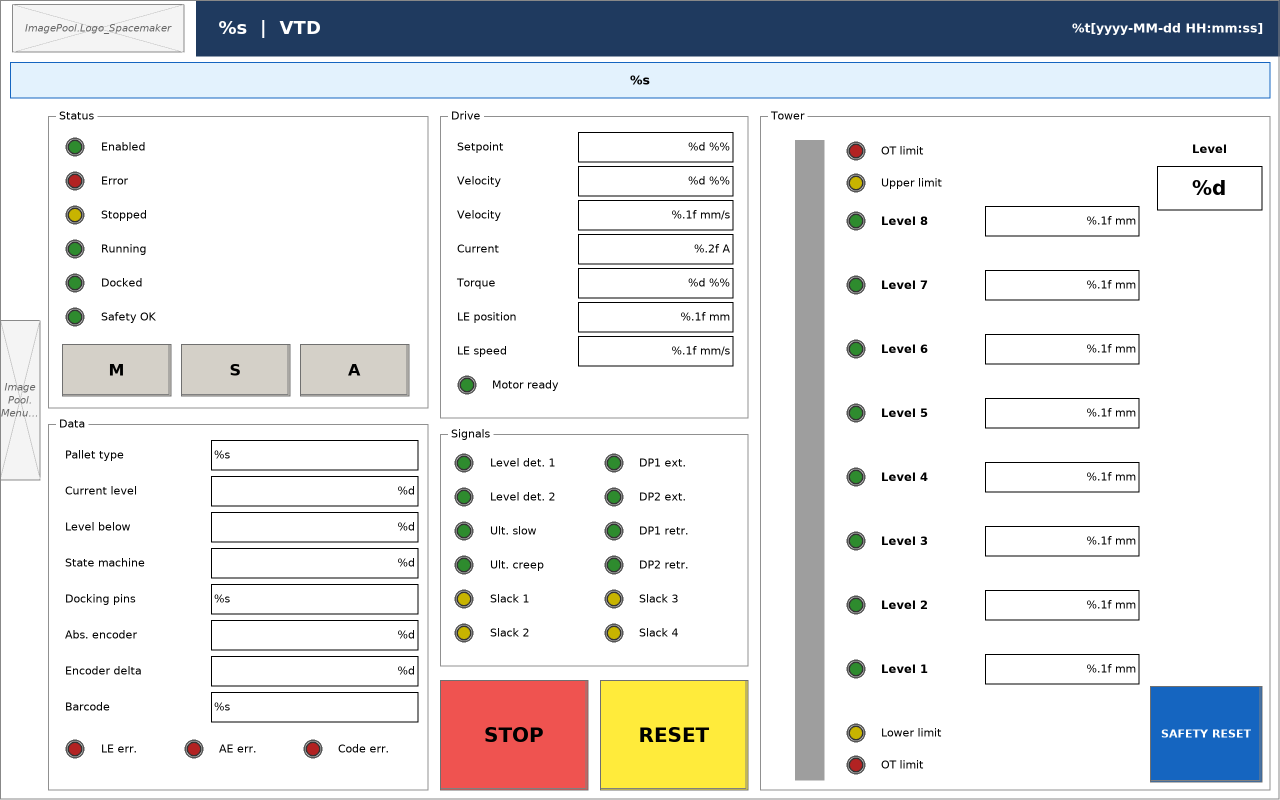
VISUALIZATION VTD  // 1280x800
    Rectangle (0,0 196x56)
        OnMouseClick: change screen: Main
    Image (12,4 172x48), image: ImagePool.Logo_Spacemaker
        OnMouseClick: change screen: Main
    Rectangle (196,0 1084x56), "%s | VTD", text variable: GVL_HMI_System.stStatus.sSystemName
    Rectangle (930,8 336x40), "%t[yyyy-MM-dd HH:mm:ss]", text variable: GVL_HMI_System.stStatus.dtNow
    Rectangle (10,62 1260x36), "%s", text variable: GVL_HMI_System.stStatus.sMessage, colour toggle: GVL_HMI_System.stStatus.bMessageAlarm
    GroupBox (48,108 380x300), "Status"
    Lamp1 (64,136 22x22), variable: GVL_HMI_VTD.stStatus.bEnabled, style: Lamp-Lamp1-Green
    Rectangle (98,132 190x30), "Enabled"
    Lamp1 (64,170 22x22), variable: GVL_HMI_VTD.stStatus.bError, style: Lamp-Lamp1-Red
    Rectangle (98,166 190x30), "Error"
    Lamp1 (64,204 22x22), variable: GVL_HMI_VTD.stStatus.bStopped, style: Lamp-Lamp1-Yellow
    Rectangle (98,200 190x30), "Stopped"
    Lamp1 (64,238 22x22), variable: GVL_HMI_VTD.stStatus.bRunning, style: Lamp-Lamp1-Green
    Rectangle (98,234 190x30), "Running"
    Lamp1 (64,272 22x22), variable: GVL_HMI_VTD.stStatus.bDocked, style: Lamp-Lamp1-Green
    Rectangle (98,268 190x30), "Docked"
    Lamp1 (64,306 22x22), variable: GVL_HMI_VTD.stStatus.bSafetyOk, style: Lamp-Lamp1-Green
    Rectangle (98,302 190x30), "Safety OK"
    Button (62,344 109x52), "M", colour toggle: GVL_HMI_VTD.stStatus.bModeManual
        tap GVL_HMI_VTD.stCommand.bModeManual p3779583253=TRUE
    Button (181,344 109x52), "S", colour toggle: GVL_HMI_VTD.stStatus.bModeSemi
        tap GVL_HMI_VTD.stCommand.bModeSemi p3779583253=TRUE
    Button (300,344 109x52), "A", colour toggle: GVL_HMI_VTD.stStatus.bModeAuto
        tap GVL_HMI_VTD.stCommand.bModeAuto p3779583253=TRUE
    GroupBox (48,416 380x374), "Data"
    Rectangle (62,440 143x30), "Pallet type"
    Rectangle (211,440 207x30), "%s", text variable: GVL_HMI_VTD.stStatus.sPalletType
    Rectangle (62,476 143x30), "Current level"
    Rectangle (211,476 207x30), "%d", text variable: GVL_HMI_VTD.stStatus.uiCurrentLevel
    Rectangle (62,512 143x30), "Level below"
    Rectangle (211,512 207x30), "%d", text variable: GVL_HMI_VTD.stStatus.uiLevelBelow
    Rectangle (62,548 143x30), "State machine"
    Rectangle (211,548 207x30), "%d", text variable: GVL_HMI_VTD.stStatus.uiStateMachine
    Rectangle (62,584 143x30), "Docking pins"
    Rectangle (211,584 207x30), "%s", text variable: GVL_HMI_VTD.stStatus.sDockingPinState
    Rectangle (62,620 143x30), "Abs. encoder"
    Rectangle (211,620 207x30), "%d", text variable: GVL_HMI_VTD.stStatus.diAbsoluteEncoder
    Rectangle (62,656 143x30), "Encoder delta"
    Rectangle (211,656 207x30), "%d", text variable: GVL_HMI_VTD.stStatus.iEncoderDelta
    Rectangle (62,692 143x30), "Barcode"
    Rectangle (211,692 207x30), "%s", text variable: GVL_HMI_VTD.stStatus.sBarcode
    Lamp1 (64,738 22x22), variable: GVL_HMI_VTD.stStatus.bLinearEncoderError, style: Lamp-Lamp1-Red
    Rectangle (98,734 78x30), "LE err."
    Lamp1 (183,738 22x22), variable: GVL_HMI_VTD.stStatus.bAbsoluteEncoderError, style: Lamp-Lamp1-Red
    Rectangle (216,734 79x30), "AE err."
    Lamp1 (302,738 22x22), variable: GVL_HMI_VTD.stStatus.bBarcodeError, style: Lamp-Lamp1-Red
    Rectangle (335,734 78x30), "Code err."
    GroupBox (440,108 308x310), "Drive"
    Rectangle (454,132 118x30), "Setpoint"
    Rectangle (578,132 155x30), "%d %%", text variable: GVL_HMI_VTD.stStatus.iSetpoint_pct
    Rectangle (454,166 118x30), "Velocity"
    Rectangle (578,166 155x30), "%d %%", text variable: GVL_HMI_VTD.stStatus.iVelocity_pct
    Rectangle (454,200 118x30), "Velocity"
    Rectangle (578,200 155x30), "%.1f mm/s", text variable: GVL_HMI_VTD.stStatus.rVelocity_mm_s
    Rectangle (454,234 118x30), "Current"
    Rectangle (578,234 155x30), "%.2f A", text variable: GVL_HMI_VTD.stStatus.rCurrent_A
    Rectangle (454,268 118x30), "Torque"
    Rectangle (578,268 155x30), "%d %%", text variable: GVL_HMI_VTD.stStatus.iTorque_pct
    Rectangle (454,302 118x30), "LE position"
    Rectangle (578,302 155x30), "%.1f mm", text variable: GVL_HMI_VTD.stStatus.rLePosition_mm
    Rectangle (454,336 118x30), "LE speed"
    Rectangle (578,336 155x30), "%.1f mm/s", text variable: GVL_HMI_VTD.stStatus.rLeSpeed_mm_s
    Lamp1 (456,374 22x22), variable: GVL_HMI_VTD.stStatus.bMotorReady, style: Lamp-Lamp1-Green
    Rectangle (489,370 190x30), "Motor ready"
    GroupBox (440,426 308x240), "Signals"
    Lamp1 (453,452 22x22), variable: GVL_HMI_VTD.stStatus.bLevelDetect1, style: Lamp-Lamp1-Green
    Rectangle (487,448 109x30), "Level det. 1"
    Lamp1 (453,486 22x22), variable: GVL_HMI_VTD.stStatus.bLevelDetect2, style: Lamp-Lamp1-Green
    Rectangle (487,482 109x30), "Level det. 2"
    Lamp1 (453,520 22x22), variable: GVL_HMI_VTD.stStatus.bUltimateSlowdown, style: Lamp-Lamp1-Green
    Rectangle (487,516 109x30), "Ult. slow"
    Lamp1 (453,554 22x22), variable: GVL_HMI_VTD.stStatus.bUltimateCreep, style: Lamp-Lamp1-Green
    Rectangle (487,550 109x30), "Ult. creep"
    Lamp1 (453,588 22x22), variable: GVL_HMI_VTD.stStatus.abChainSlack[1], style: Lamp-Lamp1-Yellow
    Rectangle (487,584 109x30), "Slack 1"
    Lamp1 (453,622 22x22), variable: GVL_HMI_VTD.stStatus.abChainSlack[2], style: Lamp-Lamp1-Yellow
    Rectangle (487,618 109x30), "Slack 2"
    Lamp1 (603,452 22x22), variable: GVL_HMI_VTD.stStatus.bDp1Extended, style: Lamp-Lamp1-Green
    Rectangle (636,448 110x30), "DP1 ext."
    Lamp1 (603,486 22x22), variable: GVL_HMI_VTD.stStatus.bDp2Extended, style: Lamp-Lamp1-Green
    Rectangle (636,482 110x30), "DP2 ext."
    Lamp1 (603,520 22x22), variable: GVL_HMI_VTD.stStatus.bDp1Retracted, style: Lamp-Lamp1-Green
    Rectangle (636,516 110x30), "DP1 retr."
    Lamp1 (603,554 22x22), variable: GVL_HMI_VTD.stStatus.bDp2Retracted, style: Lamp-Lamp1-Green
    Rectangle (636,550 110x30), "DP2 retr."
    Lamp1 (603,588 22x22), variable: GVL_HMI_VTD.stStatus.abChainSlack[3], style: Lamp-Lamp1-Yellow
    Rectangle (636,584 110x30), "Slack 3"
    Lamp1 (603,622 22x22), variable: GVL_HMI_VTD.stStatus.abChainSlack[4], style: Lamp-Lamp1-Yellow
    Rectangle (636,618 110x30), "Slack 4"
    Button (440,680 148x110), "STOP"
        tap GVL_HMI_VTD.stCommand.bStop p3779583253=TRUE
    Button (600,680 148x110), "RESET"
        tap GVL_HMI_VTD.stCommand.bReset p3779583253=TRUE
    GroupBox (760,108 510x682), "Tower"
    Rectangle (795,140 29x640)
    Lamp1 (845,140 22x22), variable: GVL_HMI_VTD.stStatus.bUpperOvertravel, style: Lamp-Lamp1-Red
    Rectangle (878,136 131x30), "OT limit"
    Lamp1 (845,172 22x22), variable: GVL_HMI_VTD.stStatus.bUpperLimit, style: Lamp-Lamp1-Yellow
    Rectangle (878,168 131x30), "Upper limit"
    Lamp1 (845,210 22x22), variable: GVL_HMI_VTD.stStatus.abLevelReached[8], style: Lamp-Lamp1-Green
    Rectangle (878,206 95x30), "Level 8"
    Rectangle (985,206 154x30), "%.1f mm", text variable: GVL_HMI_VTD.stStatus.arLevelPosition_mm[8]
    Lamp1 (845,274 22x22), variable: GVL_HMI_VTD.stStatus.abLevelReached[7], style: Lamp-Lamp1-Green
    Rectangle (878,270 95x30), "Level 7"
    Rectangle (985,270 154x30), "%.1f mm", text variable: GVL_HMI_VTD.stStatus.arLevelPosition_mm[7]
    Lamp1 (845,338 22x22), variable: GVL_HMI_VTD.stStatus.abLevelReached[6], style: Lamp-Lamp1-Green
    Rectangle (878,334 95x30), "Level 6"
    Rectangle (985,334 154x30), "%.1f mm", text variable: GVL_HMI_VTD.stStatus.arLevelPosition_mm[6]
    Lamp1 (845,402 22x22), variable: GVL_HMI_VTD.stStatus.abLevelReached[5], style: Lamp-Lamp1-Green
    Rectangle (878,398 95x30), "Level 5"
    Rectangle (985,398 154x30), "%.1f mm", text variable: GVL_HMI_VTD.stStatus.arLevelPosition_mm[5]
    Lamp1 (845,466 22x22), variable: GVL_HMI_VTD.stStatus.abLevelReached[4], style: Lamp-Lamp1-Green
    Rectangle (878,462 95x30), "Level 4"
    Rectangle (985,462 154x30), "%.1f mm", text variable: GVL_HMI_VTD.stStatus.arLevelPosition_mm[4]
    Lamp1 (845,530 22x22), variable: GVL_HMI_VTD.stStatus.abLevelReached[3], style: Lamp-Lamp1-Green
    Rectangle (878,526 95x30), "Level 3"
    Rectangle (985,526 154x30), "%.1f mm", text variable: GVL_HMI_VTD.stStatus.arLevelPosition_mm[3]
    Lamp1 (845,594 22x22), variable: GVL_HMI_VTD.stStatus.abLevelReached[2], style: Lamp-Lamp1-Green
    Rectangle (878,590 95x30), "Level 2"
    Rectangle (985,590 154x30), "%.1f mm", text variable: GVL_HMI_VTD.stStatus.arLevelPosition_mm[2]
    Lamp1 (845,658 22x22), variable: GVL_HMI_VTD.stStatus.abLevelReached[1], style: Lamp-Lamp1-Green
    Rectangle (878,654 95x30), "Level 1"
    Rectangle (985,654 154x30), "%.1f mm", text variable: GVL_HMI_VTD.stStatus.arLevelPosition_mm[1]
    Lamp1 (845,722 22x22), variable: GVL_HMI_VTD.stStatus.bLowerLimit, style: Lamp-Lamp1-Yellow
    Rectangle (878,718 131x30), "Lower limit"
    Lamp1 (845,754 22x22), variable: GVL_HMI_VTD.stStatus.bLowerOvertravel, style: Lamp-Lamp1-Red
    Rectangle (878,750 131x30), "OT limit"
    Rectangle (1157,136 105x26), "Level"
    Rectangle (1157,166 105x44), "%d", text variable: GVL_HMI_VTD.stStatus.uiCurrentLevel
    Rectangle (0,320 40x160)
        OnMouseClick: OpenDialog Dialog=Dialog, OpenModal=True, PositionX=0, PositionY=0
        OnMouseEnter: OpenDialog Dialog=Dialog, OpenModal=True, PositionX=0, PositionY=0
    Image (0,320 40x160), image: ImagePool.Menu_Tab
        OnMouseClick: OpenDialog Dialog=Dialog, OpenModal=True, PositionX=0, PositionY=0
        OnMouseEnter: OpenDialog Dialog=Dialog, OpenModal=True, PositionX=0, PositionY=0
    Button (1150,686 112x96), "SAFETY RESET", colour toggle: GVL_HMI_System.stStatus.bSafetyResetActive
        tap GVL_HMI_System.stCommand.bSafetyReset p3779583253=TRUE
END_VISUALIZATION

(* stored: Version 1.1.0.1
   Visu VTD: Id {d058b11a-4500-4a99-87d6-9345bd77b8de} *)
